(* IEC 61131-3 sources: s7-to-codesys/tests/POUs/Scenarios/FB_PumpAlternation_ScenarioTest, 7 files *)

(* ---- FB_PumpAlternation_ScenarioTest.decl.st ---- *)
// AUTO-GENERATED — не редактировать: s7conv gen-tests, сценарии scenarios/FB_PumpAlternation.csv
// Правка — в CSV (scenarios/README.md), затем python -m s7conv build-corpus.
// Назначение: тесты поведения сконвертированного FB_PumpAlternation по сценариям CSV (сценариев: 6, строк: 31):
//             один метод-тест на сценарий, строки — по порядку с моделируемым временем GVL_S7Clock.
//             Ожидаемые значения — из CSV (эталонные модели по описанию логики блока), не из
//             результата конвертации.
// Автор:      s7conv 0.1.0 (сгенерировано)
// Версия:     не указана
// Документ:   scenarios/README.md, docs/methodology.md, раздел «Проверка поведения»
FUNCTION_BLOCK FB_PumpAlternation_ScenarioTest EXTENDS coUnit.FB_TestSuite
VAR
    fbRotateOnStop : FB_PumpAlternation;  // свой экземпляр на сценарий
    xRotateOnStopDone : BOOL;  // сценарий выполнен (выполняется один раз)
    fbStandbyTakesOver : FB_PumpAlternation;  // свой экземпляр на сценарий
    xStandbyTakesOverDone : BOOL;  // сценарий выполнен (выполняется один раз)
    fbForcedAlternate : FB_PumpAlternation;  // свой экземпляр на сценарий
    xForcedAlternateDone : BOOL;  // сценарий выполнен (выполняется один раз)
    fbRotateOnStopDisabled : FB_PumpAlternation;  // свой экземпляр на сценарий
    xRotateOnStopDisabledDone : BOOL;  // сценарий выполнен (выполняется один раз)
    fbNoPumpsAvailable : FB_PumpAlternation;  // свой экземпляр на сценарий
    xNoPumpsAvailableDone : BOOL;  // сценарий выполнен (выполняется один раз)
    fbDemandClamped : FB_PumpAlternation;  // свой экземпляр на сценарий
    xDemandClampedDone : BOOL;  // сценарий выполнен (выполняется один раз)
END_VAR

(* ---- DemandClamped.method.impl.st ---- *)
// AUTO-GENERATED — не редактировать: scenarios/FB_PumpAlternation.csv, сценарий DemandClamped
coUnit.TEST('DemandClamped');
IF NOT xDemandClampedDone THEN
    xDemandClampedDone := TRUE;
    GVL_S7Clock.xSimulation := TRUE;

    // #1, t = 0 мс — demand 5 -> 3: все три
    GVL_S7Clock.tSimNow := T#0MS;
    fbDemandClamped.demand := 5;
    fbDemandClamped.available1 := TRUE;
    fbDemandClamped.available2 := TRUE;
    fbDemandClamped.available3 := TRUE;
    fbDemandClamped.alternate := FALSE;
    fbDemandClamped.rotateOnStop := TRUE;
    fbDemandClamped();
    AssertEquals_BOOL(Expected := TRUE, Actual := fbDemandClamped.run1, Message := 'DemandClamped#1 run1');
    AssertEquals_BOOL(Expected := TRUE, Actual := fbDemandClamped.run2, Message := 'DemandClamped#1 run2');
    AssertEquals_BOOL(Expected := TRUE, Actual := fbDemandClamped.run3, Message := 'DemandClamped#1 run3');
    AssertEquals_INT(Expected := 1, Actual := fbDemandClamped.leadPump, Message := 'DemandClamped#1 leadPump');
    AssertEquals_INT(Expected := 3, Actual := fbDemandClamped.runningCount, Message := 'DemandClamped#1 runningCount');
    AssertEquals_BOOL(Expected := FALSE, Actual := fbDemandClamped.shortage, Message := 'DemandClamped#1 shortage');

    // #2, t = 100 мс — demand -1 -> 0: останов, ведущий -> 2
    GVL_S7Clock.tSimNow := T#100MS;
    fbDemandClamped.demand := -1;
    fbDemandClamped();
    AssertEquals_BOOL(Expected := FALSE, Actual := fbDemandClamped.run1, Message := 'DemandClamped#2 run1');
    AssertEquals_BOOL(Expected := FALSE, Actual := fbDemandClamped.run2, Message := 'DemandClamped#2 run2');
    AssertEquals_BOOL(Expected := FALSE, Actual := fbDemandClamped.run3, Message := 'DemandClamped#2 run3');
    AssertEquals_INT(Expected := 2, Actual := fbDemandClamped.leadPump, Message := 'DemandClamped#2 leadPump');
    AssertEquals_INT(Expected := 0, Actual := fbDemandClamped.runningCount, Message := 'DemandClamped#2 runningCount');
    AssertEquals_BOOL(Expected := FALSE, Actual := fbDemandClamped.shortage, Message := 'DemandClamped#2 shortage');

    // #3, t = 200 мс — demand 4 -> 3: 2, 3, 1
    GVL_S7Clock.tSimNow := T#200MS;
    fbDemandClamped.demand := 4;
    fbDemandClamped();
    AssertEquals_BOOL(Expected := TRUE, Actual := fbDemandClamped.run1, Message := 'DemandClamped#3 run1');
    AssertEquals_BOOL(Expected := TRUE, Actual := fbDemandClamped.run2, Message := 'DemandClamped#3 run2');
    AssertEquals_BOOL(Expected := TRUE, Actual := fbDemandClamped.run3, Message := 'DemandClamped#3 run3');
    AssertEquals_INT(Expected := 2, Actual := fbDemandClamped.leadPump, Message := 'DemandClamped#3 leadPump');
    AssertEquals_INT(Expected := 3, Actual := fbDemandClamped.runningCount, Message := 'DemandClamped#3 runningCount');
    AssertEquals_BOOL(Expected := FALSE, Actual := fbDemandClamped.shortage, Message := 'DemandClamped#3 shortage');

    GVL_S7Clock.xSimulation := FALSE;
END_IF
coUnit.TEST_FINISHED();

(* ---- ForcedAlternate.method.impl.st ---- *)
// AUTO-GENERATED — не редактировать: scenarios/FB_PumpAlternation.csv, сценарий ForcedAlternate
coUnit.TEST('ForcedAlternate');
IF NOT xForcedAlternateDone THEN
    xForcedAlternateDone := TRUE;
    GVL_S7Clock.xSimulation := TRUE;

    // #1, t = 0 мс — один насос: 1
    GVL_S7Clock.tSimNow := T#0MS;
    fbForcedAlternate.demand := 1;
    fbForcedAlternate.available1 := TRUE;
    fbForcedAlternate.available2 := TRUE;
    fbForcedAlternate.available3 := TRUE;
    fbForcedAlternate.alternate := FALSE;
    fbForcedAlternate.rotateOnStop := TRUE;
    fbForcedAlternate();
    AssertEquals_BOOL(Expected := TRUE, Actual := fbForcedAlternate.run1, Message := 'ForcedAlternate#1 run1');
    AssertEquals_BOOL(Expected := FALSE, Actual := fbForcedAlternate.run2, Message := 'ForcedAlternate#1 run2');
    AssertEquals_BOOL(Expected := FALSE, Actual := fbForcedAlternate.run3, Message := 'ForcedAlternate#1 run3');
    AssertEquals_INT(Expected := 1, Actual := fbForcedAlternate.leadPump, Message := 'ForcedAlternate#1 leadPump');
    AssertEquals_INT(Expected := 1,
                     Actual := fbForcedAlternate.runningCount,
                     Message := 'ForcedAlternate#1 runningCount');
    AssertEquals_BOOL(Expected := FALSE, Actual := fbForcedAlternate.shortage, Message := 'ForcedAlternate#1 shortage');

    // #2, t = 100 мс — фронт alternate: ведущий 2, переключение в работе
    GVL_S7Clock.tSimNow := T#100MS;
    fbForcedAlternate.alternate := TRUE;
    fbForcedAlternate();
    AssertEquals_BOOL(Expected := FALSE, Actual := fbForcedAlternate.run1, Message := 'ForcedAlternate#2 run1');
    AssertEquals_BOOL(Expected := TRUE, Actual := fbForcedAlternate.run2, Message := 'ForcedAlternate#2 run2');
    AssertEquals_BOOL(Expected := FALSE, Actual := fbForcedAlternate.run3, Message := 'ForcedAlternate#2 run3');
    AssertEquals_INT(Expected := 2, Actual := fbForcedAlternate.leadPump, Message := 'ForcedAlternate#2 leadPump');
    AssertEquals_INT(Expected := 1,
                     Actual := fbForcedAlternate.runningCount,
                     Message := 'ForcedAlternate#2 runningCount');
    AssertEquals_BOOL(Expected := FALSE, Actual := fbForcedAlternate.shortage, Message := 'ForcedAlternate#2 shortage');

    // #3, t = 200 мс — alternate держится: фронта нет
    GVL_S7Clock.tSimNow := T#200MS;
    fbForcedAlternate();
    AssertEquals_BOOL(Expected := FALSE, Actual := fbForcedAlternate.run1, Message := 'ForcedAlternate#3 run1');
    AssertEquals_BOOL(Expected := TRUE, Actual := fbForcedAlternate.run2, Message := 'ForcedAlternate#3 run2');
    AssertEquals_BOOL(Expected := FALSE, Actual := fbForcedAlternate.run3, Message := 'ForcedAlternate#3 run3');
    AssertEquals_INT(Expected := 2, Actual := fbForcedAlternate.leadPump, Message := 'ForcedAlternate#3 leadPump');
    AssertEquals_INT(Expected := 1,
                     Actual := fbForcedAlternate.runningCount,
                     Message := 'ForcedAlternate#3 runningCount');
    AssertEquals_BOOL(Expected := FALSE, Actual := fbForcedAlternate.shortage, Message := 'ForcedAlternate#3 shortage');

    // #4, t = 300 мс — отпущен
    GVL_S7Clock.tSimNow := T#300MS;
    fbForcedAlternate.alternate := FALSE;
    fbForcedAlternate();
    AssertEquals_BOOL(Expected := FALSE, Actual := fbForcedAlternate.run1, Message := 'ForcedAlternate#4 run1');
    AssertEquals_BOOL(Expected := TRUE, Actual := fbForcedAlternate.run2, Message := 'ForcedAlternate#4 run2');
    AssertEquals_BOOL(Expected := FALSE, Actual := fbForcedAlternate.run3, Message := 'ForcedAlternate#4 run3');
    AssertEquals_INT(Expected := 2, Actual := fbForcedAlternate.leadPump, Message := 'ForcedAlternate#4 leadPump');
    AssertEquals_INT(Expected := 1,
                     Actual := fbForcedAlternate.runningCount,
                     Message := 'ForcedAlternate#4 runningCount');
    AssertEquals_BOOL(Expected := FALSE, Actual := fbForcedAlternate.shortage, Message := 'ForcedAlternate#4 shortage');

    // #5, t = 400 мс — фронт: ведущий 3
    GVL_S7Clock.tSimNow := T#400MS;
    fbForcedAlternate.alternate := TRUE;
    fbForcedAlternate();
    AssertEquals_BOOL(Expected := FALSE, Actual := fbForcedAlternate.run1, Message := 'ForcedAlternate#5 run1');
    AssertEquals_BOOL(Expected := FALSE, Actual := fbForcedAlternate.run2, Message := 'ForcedAlternate#5 run2');
    AssertEquals_BOOL(Expected := TRUE, Actual := fbForcedAlternate.run3, Message := 'ForcedAlternate#5 run3');
    AssertEquals_INT(Expected := 3, Actual := fbForcedAlternate.leadPump, Message := 'ForcedAlternate#5 leadPump');
    AssertEquals_INT(Expected := 1,
                     Actual := fbForcedAlternate.runningCount,
                     Message := 'ForcedAlternate#5 runningCount');
    AssertEquals_BOOL(Expected := FALSE, Actual := fbForcedAlternate.shortage, Message := 'ForcedAlternate#5 shortage');

    GVL_S7Clock.xSimulation := FALSE;
END_IF
coUnit.TEST_FINISHED();

(* ---- NoPumpsAvailable.method.impl.st ---- *)
// AUTO-GENERATED — не редактировать: scenarios/FB_PumpAlternation.csv, сценарий NoPumpsAvailable
coUnit.TEST('NoPumpsAvailable');
IF NOT xNoPumpsAvailableDone THEN
    xNoPumpsAvailableDone := TRUE;
    GVL_S7Clock.xSimulation := TRUE;

    // #1, t = 0 мс — нужно 2, доступных нет: нехватка
    GVL_S7Clock.tSimNow := T#0MS;
    fbNoPumpsAvailable.demand := 2;
    fbNoPumpsAvailable.available1 := FALSE;
    fbNoPumpsAvailable.available2 := FALSE;
    fbNoPumpsAvailable.available3 := FALSE;
    fbNoPumpsAvailable.alternate := FALSE;
    fbNoPumpsAvailable.rotateOnStop := TRUE;
    fbNoPumpsAvailable();
    AssertEquals_BOOL(Expected := FALSE, Actual := fbNoPumpsAvailable.run1, Message := 'NoPumpsAvailable#1 run1');
    AssertEquals_BOOL(Expected := FALSE, Actual := fbNoPumpsAvailable.run2, Message := 'NoPumpsAvailable#1 run2');
    AssertEquals_BOOL(Expected := FALSE, Actual := fbNoPumpsAvailable.run3, Message := 'NoPumpsAvailable#1 run3');
    AssertEquals_INT(Expected := 1, Actual := fbNoPumpsAvailable.leadPump, Message := 'NoPumpsAvailable#1 leadPump');
    AssertEquals_INT(Expected := 0,
                     Actual := fbNoPumpsAvailable.runningCount,
                     Message := 'NoPumpsAvailable#1 runningCount');
    AssertEquals_BOOL(Expected := TRUE,
                      Actual := fbNoPumpsAvailable.shortage,
                      Message := 'NoPumpsAvailable#1 shortage');

    // #2, t = 100 мс — останов: искать некого, ведущий 1
    GVL_S7Clock.tSimNow := T#100MS;
    fbNoPumpsAvailable.demand := 0;
    fbNoPumpsAvailable();
    AssertEquals_BOOL(Expected := FALSE, Actual := fbNoPumpsAvailable.run1, Message := 'NoPumpsAvailable#2 run1');
    AssertEquals_BOOL(Expected := FALSE, Actual := fbNoPumpsAvailable.run2, Message := 'NoPumpsAvailable#2 run2');
    AssertEquals_BOOL(Expected := FALSE, Actual := fbNoPumpsAvailable.run3, Message := 'NoPumpsAvailable#2 run3');
    AssertEquals_INT(Expected := 1, Actual := fbNoPumpsAvailable.leadPump, Message := 'NoPumpsAvailable#2 leadPump');
    AssertEquals_INT(Expected := 0,
                     Actual := fbNoPumpsAvailable.runningCount,
                     Message := 'NoPumpsAvailable#2 runningCount');
    AssertEquals_BOOL(Expected := FALSE,
                      Actual := fbNoPumpsAvailable.shortage,
                      Message := 'NoPumpsAvailable#2 shortage');

    // #3, t = 200 мс — фронт alternate: искать некого, ведущий 1
    GVL_S7Clock.tSimNow := T#200MS;
    fbNoPumpsAvailable.alternate := TRUE;
    fbNoPumpsAvailable();
    AssertEquals_BOOL(Expected := FALSE, Actual := fbNoPumpsAvailable.run1, Message := 'NoPumpsAvailable#3 run1');
    AssertEquals_BOOL(Expected := FALSE, Actual := fbNoPumpsAvailable.run2, Message := 'NoPumpsAvailable#3 run2');
    AssertEquals_BOOL(Expected := FALSE, Actual := fbNoPumpsAvailable.run3, Message := 'NoPumpsAvailable#3 run3');
    AssertEquals_INT(Expected := 1, Actual := fbNoPumpsAvailable.leadPump, Message := 'NoPumpsAvailable#3 leadPump');
    AssertEquals_INT(Expected := 0,
                     Actual := fbNoPumpsAvailable.runningCount,
                     Message := 'NoPumpsAvailable#3 runningCount');
    AssertEquals_BOOL(Expected := FALSE,
                      Actual := fbNoPumpsAvailable.shortage,
                      Message := 'NoPumpsAvailable#3 shortage');

    // #4, t = 300 мс — доступен только 3: работает 3, ведущий 1
    GVL_S7Clock.tSimNow := T#300MS;
    fbNoPumpsAvailable.demand := 1;
    fbNoPumpsAvailable.available3 := TRUE;
    fbNoPumpsAvailable.alternate := FALSE;
    fbNoPumpsAvailable();
    AssertEquals_BOOL(Expected := FALSE, Actual := fbNoPumpsAvailable.run1, Message := 'NoPumpsAvailable#4 run1');
    AssertEquals_BOOL(Expected := FALSE, Actual := fbNoPumpsAvailable.run2, Message := 'NoPumpsAvailable#4 run2');
    AssertEquals_BOOL(Expected := TRUE, Actual := fbNoPumpsAvailable.run3, Message := 'NoPumpsAvailable#4 run3');
    AssertEquals_INT(Expected := 1, Actual := fbNoPumpsAvailable.leadPump, Message := 'NoPumpsAvailable#4 leadPump');
    AssertEquals_INT(Expected := 1,
                     Actual := fbNoPumpsAvailable.runningCount,
                     Message := 'NoPumpsAvailable#4 runningCount');
    AssertEquals_BOOL(Expected := FALSE,
                      Actual := fbNoPumpsAvailable.shortage,
                      Message := 'NoPumpsAvailable#4 shortage');

    GVL_S7Clock.xSimulation := FALSE;
END_IF
coUnit.TEST_FINISHED();

(* ---- RotateOnStop.method.impl.st ---- *)
// AUTO-GENERATED — не редактировать: scenarios/FB_PumpAlternation.csv, сценарий RotateOnStop
coUnit.TEST('RotateOnStop');
IF NOT xRotateOnStopDone THEN
    xRotateOnStopDone := TRUE;
    GVL_S7Clock.xSimulation := TRUE;

    // #1, t = 0 мс — первый вызов при demand = 0: спада нет, ведущий 1
    GVL_S7Clock.tSimNow := T#0MS;
    fbRotateOnStop.demand := 0;
    fbRotateOnStop.available1 := TRUE;
    fbRotateOnStop.available2 := TRUE;
    fbRotateOnStop.available3 := TRUE;
    fbRotateOnStop.alternate := FALSE;
    fbRotateOnStop.rotateOnStop := TRUE;
    fbRotateOnStop();
    AssertEquals_BOOL(Expected := FALSE, Actual := fbRotateOnStop.run1, Message := 'RotateOnStop#1 run1');
    AssertEquals_BOOL(Expected := FALSE, Actual := fbRotateOnStop.run2, Message := 'RotateOnStop#1 run2');
    AssertEquals_BOOL(Expected := FALSE, Actual := fbRotateOnStop.run3, Message := 'RotateOnStop#1 run3');
    AssertEquals_INT(Expected := 1, Actual := fbRotateOnStop.leadPump, Message := 'RotateOnStop#1 leadPump');
    AssertEquals_INT(Expected := 0, Actual := fbRotateOnStop.runningCount, Message := 'RotateOnStop#1 runningCount');
    AssertEquals_BOOL(Expected := FALSE, Actual := fbRotateOnStop.shortage, Message := 'RotateOnStop#1 shortage');

    // #2, t = 100 мс — один насос: ведущий 1
    GVL_S7Clock.tSimNow := T#100MS;
    fbRotateOnStop.demand := 1;
    fbRotateOnStop();
    AssertEquals_BOOL(Expected := TRUE, Actual := fbRotateOnStop.run1, Message := 'RotateOnStop#2 run1');
    AssertEquals_BOOL(Expected := FALSE, Actual := fbRotateOnStop.run2, Message := 'RotateOnStop#2 run2');
    AssertEquals_BOOL(Expected := FALSE, Actual := fbRotateOnStop.run3, Message := 'RotateOnStop#2 run3');
    AssertEquals_INT(Expected := 1, Actual := fbRotateOnStop.leadPump, Message := 'RotateOnStop#2 leadPump');
    AssertEquals_INT(Expected := 1, Actual := fbRotateOnStop.runningCount, Message := 'RotateOnStop#2 runningCount');
    AssertEquals_BOOL(Expected := FALSE, Actual := fbRotateOnStop.shortage, Message := 'RotateOnStop#2 shortage');

    // #3, t = 200 мс — два насоса: 1 и 2
    GVL_S7Clock.tSimNow := T#200MS;
    fbRotateOnStop.demand := 2;
    fbRotateOnStop();
    AssertEquals_BOOL(Expected := TRUE, Actual := fbRotateOnStop.run1, Message := 'RotateOnStop#3 run1');
    AssertEquals_BOOL(Expected := TRUE, Actual := fbRotateOnStop.run2, Message := 'RotateOnStop#3 run2');
    AssertEquals_BOOL(Expected := FALSE, Actual := fbRotateOnStop.run3, Message := 'RotateOnStop#3 run3');
    AssertEquals_INT(Expected := 1, Actual := fbRotateOnStop.leadPump, Message := 'RotateOnStop#3 leadPump');
    AssertEquals_INT(Expected := 2, Actual := fbRotateOnStop.runningCount, Message := 'RotateOnStop#3 runningCount');
    AssertEquals_BOOL(Expected := FALSE, Actual := fbRotateOnStop.shortage, Message := 'RotateOnStop#3 shortage');

    // #4, t = 300 мс — останов группы: ведущий -> 2
    GVL_S7Clock.tSimNow := T#300MS;
    fbRotateOnStop.demand := 0;
    fbRotateOnStop();
    AssertEquals_BOOL(Expected := FALSE, Actual := fbRotateOnStop.run1, Message := 'RotateOnStop#4 run1');
    AssertEquals_BOOL(Expected := FALSE, Actual := fbRotateOnStop.run2, Message := 'RotateOnStop#4 run2');
    AssertEquals_BOOL(Expected := FALSE, Actual := fbRotateOnStop.run3, Message := 'RotateOnStop#4 run3');
    AssertEquals_INT(Expected := 2, Actual := fbRotateOnStop.leadPump, Message := 'RotateOnStop#4 leadPump');
    AssertEquals_INT(Expected := 0, Actual := fbRotateOnStop.runningCount, Message := 'RotateOnStop#4 runningCount');
    AssertEquals_BOOL(Expected := FALSE, Actual := fbRotateOnStop.shortage, Message := 'RotateOnStop#4 shortage');

    // #5, t = 400 мс — один насос: 2
    GVL_S7Clock.tSimNow := T#400MS;
    fbRotateOnStop.demand := 1;
    fbRotateOnStop();
    AssertEquals_BOOL(Expected := FALSE, Actual := fbRotateOnStop.run1, Message := 'RotateOnStop#5 run1');
    AssertEquals_BOOL(Expected := TRUE, Actual := fbRotateOnStop.run2, Message := 'RotateOnStop#5 run2');
    AssertEquals_BOOL(Expected := FALSE, Actual := fbRotateOnStop.run3, Message := 'RotateOnStop#5 run3');
    AssertEquals_INT(Expected := 2, Actual := fbRotateOnStop.leadPump, Message := 'RotateOnStop#5 leadPump');
    AssertEquals_INT(Expected := 1, Actual := fbRotateOnStop.runningCount, Message := 'RotateOnStop#5 runningCount');
    AssertEquals_BOOL(Expected := FALSE, Actual := fbRotateOnStop.shortage, Message := 'RotateOnStop#5 shortage');

    // #6, t = 500 мс — три насоса: 2, 3, 1
    GVL_S7Clock.tSimNow := T#500MS;
    fbRotateOnStop.demand := 3;
    fbRotateOnStop();
    AssertEquals_BOOL(Expected := TRUE, Actual := fbRotateOnStop.run1, Message := 'RotateOnStop#6 run1');
    AssertEquals_BOOL(Expected := TRUE, Actual := fbRotateOnStop.run2, Message := 'RotateOnStop#6 run2');
    AssertEquals_BOOL(Expected := TRUE, Actual := fbRotateOnStop.run3, Message := 'RotateOnStop#6 run3');
    AssertEquals_INT(Expected := 2, Actual := fbRotateOnStop.leadPump, Message := 'RotateOnStop#6 leadPump');
    AssertEquals_INT(Expected := 3, Actual := fbRotateOnStop.runningCount, Message := 'RotateOnStop#6 runningCount');
    AssertEquals_BOOL(Expected := FALSE, Actual := fbRotateOnStop.shortage, Message := 'RotateOnStop#6 shortage');

    // #7, t = 600 мс — останов: ведущий -> 3
    GVL_S7Clock.tSimNow := T#600MS;
    fbRotateOnStop.demand := 0;
    fbRotateOnStop();
    AssertEquals_BOOL(Expected := FALSE, Actual := fbRotateOnStop.run1, Message := 'RotateOnStop#7 run1');
    AssertEquals_BOOL(Expected := FALSE, Actual := fbRotateOnStop.run2, Message := 'RotateOnStop#7 run2');
    AssertEquals_BOOL(Expected := FALSE, Actual := fbRotateOnStop.run3, Message := 'RotateOnStop#7 run3');
    AssertEquals_INT(Expected := 3, Actual := fbRotateOnStop.leadPump, Message := 'RotateOnStop#7 leadPump');
    AssertEquals_INT(Expected := 0, Actual := fbRotateOnStop.runningCount, Message := 'RotateOnStop#7 runningCount');
    AssertEquals_BOOL(Expected := FALSE, Actual := fbRotateOnStop.shortage, Message := 'RotateOnStop#7 shortage');

    // #8, t = 700 мс — один насос: 3
    GVL_S7Clock.tSimNow := T#700MS;
    fbRotateOnStop.demand := 1;
    fbRotateOnStop();
    AssertEquals_BOOL(Expected := FALSE, Actual := fbRotateOnStop.run1, Message := 'RotateOnStop#8 run1');
    AssertEquals_BOOL(Expected := FALSE, Actual := fbRotateOnStop.run2, Message := 'RotateOnStop#8 run2');
    AssertEquals_BOOL(Expected := TRUE, Actual := fbRotateOnStop.run3, Message := 'RotateOnStop#8 run3');
    AssertEquals_INT(Expected := 3, Actual := fbRotateOnStop.leadPump, Message := 'RotateOnStop#8 leadPump');
    AssertEquals_INT(Expected := 1, Actual := fbRotateOnStop.runningCount, Message := 'RotateOnStop#8 runningCount');
    AssertEquals_BOOL(Expected := FALSE, Actual := fbRotateOnStop.shortage, Message := 'RotateOnStop#8 shortage');

    // #9, t = 800 мс — останов: ведущий -> 1 (по кругу)
    GVL_S7Clock.tSimNow := T#800MS;
    fbRotateOnStop.demand := 0;
    fbRotateOnStop();
    AssertEquals_BOOL(Expected := FALSE, Actual := fbRotateOnStop.run1, Message := 'RotateOnStop#9 run1');
    AssertEquals_BOOL(Expected := FALSE, Actual := fbRotateOnStop.run2, Message := 'RotateOnStop#9 run2');
    AssertEquals_BOOL(Expected := FALSE, Actual := fbRotateOnStop.run3, Message := 'RotateOnStop#9 run3');
    AssertEquals_INT(Expected := 1, Actual := fbRotateOnStop.leadPump, Message := 'RotateOnStop#9 leadPump');
    AssertEquals_INT(Expected := 0, Actual := fbRotateOnStop.runningCount, Message := 'RotateOnStop#9 runningCount');
    AssertEquals_BOOL(Expected := FALSE, Actual := fbRotateOnStop.shortage, Message := 'RotateOnStop#9 shortage');

    // #10, t = 900 мс — demand остаётся 0: спада нет, ведущий 1
    GVL_S7Clock.tSimNow := T#900MS;
    fbRotateOnStop();
    AssertEquals_BOOL(Expected := FALSE, Actual := fbRotateOnStop.run1, Message := 'RotateOnStop#10 run1');
    AssertEquals_BOOL(Expected := FALSE, Actual := fbRotateOnStop.run2, Message := 'RotateOnStop#10 run2');
    AssertEquals_BOOL(Expected := FALSE, Actual := fbRotateOnStop.run3, Message := 'RotateOnStop#10 run3');
    AssertEquals_INT(Expected := 1, Actual := fbRotateOnStop.leadPump, Message := 'RotateOnStop#10 leadPump');
    AssertEquals_INT(Expected := 0, Actual := fbRotateOnStop.runningCount, Message := 'RotateOnStop#10 runningCount');
    AssertEquals_BOOL(Expected := FALSE, Actual := fbRotateOnStop.shortage, Message := 'RotateOnStop#10 shortage');

    GVL_S7Clock.xSimulation := FALSE;
END_IF
coUnit.TEST_FINISHED();

(* ---- RotateOnStopDisabled.method.impl.st ---- *)
// AUTO-GENERATED — не редактировать: scenarios/FB_PumpAlternation.csv, сценарий RotateOnStopDisabled
coUnit.TEST('RotateOnStopDisabled');
IF NOT xRotateOnStopDisabledDone THEN
    xRotateOnStopDisabledDone := TRUE;
    GVL_S7Clock.xSimulation := TRUE;

    // #1, t = 0 мс — один насос: 1
    GVL_S7Clock.tSimNow := T#0MS;
    fbRotateOnStopDisabled.demand := 1;
    fbRotateOnStopDisabled.available1 := TRUE;
    fbRotateOnStopDisabled.available2 := TRUE;
    fbRotateOnStopDisabled.available3 := TRUE;
    fbRotateOnStopDisabled.alternate := FALSE;
    fbRotateOnStopDisabled.rotateOnStop := FALSE;
    fbRotateOnStopDisabled();
    AssertEquals_BOOL(Expected := TRUE,
                      Actual := fbRotateOnStopDisabled.run1,
                      Message := 'RotateOnStopDisabled#1 run1');
    AssertEquals_BOOL(Expected := FALSE,
                      Actual := fbRotateOnStopDisabled.run2,
                      Message := 'RotateOnStopDisabled#1 run2');
    AssertEquals_BOOL(Expected := FALSE,
                      Actual := fbRotateOnStopDisabled.run3,
                      Message := 'RotateOnStopDisabled#1 run3');
    AssertEquals_INT(Expected := 1,
                     Actual := fbRotateOnStopDisabled.leadPump,
                     Message := 'RotateOnStopDisabled#1 leadPump');
    AssertEquals_INT(Expected := 1,
                     Actual := fbRotateOnStopDisabled.runningCount,
                     Message := 'RotateOnStopDisabled#1 runningCount');
    AssertEquals_BOOL(Expected := FALSE,
                      Actual := fbRotateOnStopDisabled.shortage,
                      Message := 'RotateOnStopDisabled#1 shortage');

    // #2, t = 100 мс — останов: ведущий остаётся 1
    GVL_S7Clock.tSimNow := T#100MS;
    fbRotateOnStopDisabled.demand := 0;
    fbRotateOnStopDisabled();
    AssertEquals_BOOL(Expected := FALSE,
                      Actual := fbRotateOnStopDisabled.run1,
                      Message := 'RotateOnStopDisabled#2 run1');
    AssertEquals_BOOL(Expected := FALSE,
                      Actual := fbRotateOnStopDisabled.run2,
                      Message := 'RotateOnStopDisabled#2 run2');
    AssertEquals_BOOL(Expected := FALSE,
                      Actual := fbRotateOnStopDisabled.run3,
                      Message := 'RotateOnStopDisabled#2 run3');
    AssertEquals_INT(Expected := 1,
                     Actual := fbRotateOnStopDisabled.leadPump,
                     Message := 'RotateOnStopDisabled#2 leadPump');
    AssertEquals_INT(Expected := 0,
                     Actual := fbRotateOnStopDisabled.runningCount,
                     Message := 'RotateOnStopDisabled#2 runningCount');
    AssertEquals_BOOL(Expected := FALSE,
                      Actual := fbRotateOnStopDisabled.shortage,
                      Message := 'RotateOnStopDisabled#2 shortage');

    // #3, t = 200 мс — снова 1
    GVL_S7Clock.tSimNow := T#200MS;
    fbRotateOnStopDisabled.demand := 1;
    fbRotateOnStopDisabled();
    AssertEquals_BOOL(Expected := TRUE,
                      Actual := fbRotateOnStopDisabled.run1,
                      Message := 'RotateOnStopDisabled#3 run1');
    AssertEquals_BOOL(Expected := FALSE,
                      Actual := fbRotateOnStopDisabled.run2,
                      Message := 'RotateOnStopDisabled#3 run2');
    AssertEquals_BOOL(Expected := FALSE,
                      Actual := fbRotateOnStopDisabled.run3,
                      Message := 'RotateOnStopDisabled#3 run3');
    AssertEquals_INT(Expected := 1,
                     Actual := fbRotateOnStopDisabled.leadPump,
                     Message := 'RotateOnStopDisabled#3 leadPump');
    AssertEquals_INT(Expected := 1,
                     Actual := fbRotateOnStopDisabled.runningCount,
                     Message := 'RotateOnStopDisabled#3 runningCount');
    AssertEquals_BOOL(Expected := FALSE,
                      Actual := fbRotateOnStopDisabled.shortage,
                      Message := 'RotateOnStopDisabled#3 shortage');

    GVL_S7Clock.xSimulation := FALSE;
END_IF
coUnit.TEST_FINISHED();

(* ---- StandbyTakesOver.method.impl.st ---- *)
// AUTO-GENERATED — не редактировать: scenarios/FB_PumpAlternation.csv, сценарий StandbyTakesOver
coUnit.TEST('StandbyTakesOver');
IF NOT xStandbyTakesOverDone THEN
    xStandbyTakesOverDone := TRUE;
    GVL_S7Clock.xSimulation := TRUE;

    // #1, t = 0 мс — один насос: 1
    GVL_S7Clock.tSimNow := T#0MS;
    fbStandbyTakesOver.demand := 1;
    fbStandbyTakesOver.available1 := TRUE;
    fbStandbyTakesOver.available2 := TRUE;
    fbStandbyTakesOver.available3 := TRUE;
    fbStandbyTakesOver.alternate := FALSE;
    fbStandbyTakesOver.rotateOnStop := TRUE;
    fbStandbyTakesOver();
    AssertEquals_BOOL(Expected := TRUE, Actual := fbStandbyTakesOver.run1, Message := 'StandbyTakesOver#1 run1');
    AssertEquals_BOOL(Expected := FALSE, Actual := fbStandbyTakesOver.run2, Message := 'StandbyTakesOver#1 run2');
    AssertEquals_BOOL(Expected := FALSE, Actual := fbStandbyTakesOver.run3, Message := 'StandbyTakesOver#1 run3');
    AssertEquals_INT(Expected := 1, Actual := fbStandbyTakesOver.leadPump, Message := 'StandbyTakesOver#1 leadPump');
    AssertEquals_INT(Expected := 1,
                     Actual := fbStandbyTakesOver.runningCount,
                     Message := 'StandbyTakesOver#1 runningCount');
    AssertEquals_BOOL(Expected := FALSE,
                      Actual := fbStandbyTakesOver.shortage,
                      Message := 'StandbyTakesOver#1 shortage');

    // #2, t = 100 мс — насос 1 недоступен: работает 2, ведущий остаётся 1
    GVL_S7Clock.tSimNow := T#100MS;
    fbStandbyTakesOver.available1 := FALSE;
    fbStandbyTakesOver();
    AssertEquals_BOOL(Expected := FALSE, Actual := fbStandbyTakesOver.run1, Message := 'StandbyTakesOver#2 run1');
    AssertEquals_BOOL(Expected := TRUE, Actual := fbStandbyTakesOver.run2, Message := 'StandbyTakesOver#2 run2');
    AssertEquals_BOOL(Expected := FALSE, Actual := fbStandbyTakesOver.run3, Message := 'StandbyTakesOver#2 run3');
    AssertEquals_INT(Expected := 1, Actual := fbStandbyTakesOver.leadPump, Message := 'StandbyTakesOver#2 leadPump');
    AssertEquals_INT(Expected := 1,
                     Actual := fbStandbyTakesOver.runningCount,
                     Message := 'StandbyTakesOver#2 runningCount');
    AssertEquals_BOOL(Expected := FALSE,
                      Actual := fbStandbyTakesOver.shortage,
                      Message := 'StandbyTakesOver#2 shortage');

    // #3, t = 200 мс — насос 1 вернулся: снова 1
    GVL_S7Clock.tSimNow := T#200MS;
    fbStandbyTakesOver.available1 := TRUE;
    fbStandbyTakesOver();
    AssertEquals_BOOL(Expected := TRUE, Actual := fbStandbyTakesOver.run1, Message := 'StandbyTakesOver#3 run1');
    AssertEquals_BOOL(Expected := FALSE, Actual := fbStandbyTakesOver.run2, Message := 'StandbyTakesOver#3 run2');
    AssertEquals_BOOL(Expected := FALSE, Actual := fbStandbyTakesOver.run3, Message := 'StandbyTakesOver#3 run3');
    AssertEquals_INT(Expected := 1, Actual := fbStandbyTakesOver.leadPump, Message := 'StandbyTakesOver#3 leadPump');
    AssertEquals_INT(Expected := 1,
                     Actual := fbStandbyTakesOver.runningCount,
                     Message := 'StandbyTakesOver#3 runningCount');
    AssertEquals_BOOL(Expected := FALSE,
                      Actual := fbStandbyTakesOver.shortage,
                      Message := 'StandbyTakesOver#3 shortage');

    // #4, t = 300 мс — нужно 3, доступно 2: 1 и 3, нехватка
    GVL_S7Clock.tSimNow := T#300MS;
    fbStandbyTakesOver.demand := 3;
    fbStandbyTakesOver.available2 := FALSE;
    fbStandbyTakesOver();
    AssertEquals_BOOL(Expected := TRUE, Actual := fbStandbyTakesOver.run1, Message := 'StandbyTakesOver#4 run1');
    AssertEquals_BOOL(Expected := FALSE, Actual := fbStandbyTakesOver.run2, Message := 'StandbyTakesOver#4 run2');
    AssertEquals_BOOL(Expected := TRUE, Actual := fbStandbyTakesOver.run3, Message := 'StandbyTakesOver#4 run3');
    AssertEquals_INT(Expected := 1, Actual := fbStandbyTakesOver.leadPump, Message := 'StandbyTakesOver#4 leadPump');
    AssertEquals_INT(Expected := 2,
                     Actual := fbStandbyTakesOver.runningCount,
                     Message := 'StandbyTakesOver#4 runningCount');
    AssertEquals_BOOL(Expected := TRUE,
                      Actual := fbStandbyTakesOver.shortage,
                      Message := 'StandbyTakesOver#4 shortage');

    // #5, t = 400 мс — останов: после 1 недоступен 2 — ведущий 3
    GVL_S7Clock.tSimNow := T#400MS;
    fbStandbyTakesOver.demand := 0;
    fbStandbyTakesOver();
    AssertEquals_BOOL(Expected := FALSE, Actual := fbStandbyTakesOver.run1, Message := 'StandbyTakesOver#5 run1');
    AssertEquals_BOOL(Expected := FALSE, Actual := fbStandbyTakesOver.run2, Message := 'StandbyTakesOver#5 run2');
    AssertEquals_BOOL(Expected := FALSE, Actual := fbStandbyTakesOver.run3, Message := 'StandbyTakesOver#5 run3');
    AssertEquals_INT(Expected := 3, Actual := fbStandbyTakesOver.leadPump, Message := 'StandbyTakesOver#5 leadPump');
    AssertEquals_INT(Expected := 0,
                     Actual := fbStandbyTakesOver.runningCount,
                     Message := 'StandbyTakesOver#5 runningCount');
    AssertEquals_BOOL(Expected := FALSE,
                      Actual := fbStandbyTakesOver.shortage,
                      Message := 'StandbyTakesOver#5 shortage');

    // #6, t = 500 мс — один насос: 3
    GVL_S7Clock.tSimNow := T#500MS;
    fbStandbyTakesOver.demand := 1;
    fbStandbyTakesOver();
    AssertEquals_BOOL(Expected := FALSE, Actual := fbStandbyTakesOver.run1, Message := 'StandbyTakesOver#6 run1');
    AssertEquals_BOOL(Expected := FALSE, Actual := fbStandbyTakesOver.run2, Message := 'StandbyTakesOver#6 run2');
    AssertEquals_BOOL(Expected := TRUE, Actual := fbStandbyTakesOver.run3, Message := 'StandbyTakesOver#6 run3');
    AssertEquals_INT(Expected := 3, Actual := fbStandbyTakesOver.leadPump, Message := 'StandbyTakesOver#6 leadPump');
    AssertEquals_INT(Expected := 1,
                     Actual := fbStandbyTakesOver.runningCount,
                     Message := 'StandbyTakesOver#6 runningCount');
    AssertEquals_BOOL(Expected := FALSE,
                      Actual := fbStandbyTakesOver.shortage,
                      Message := 'StandbyTakesOver#6 shortage');

    GVL_S7Clock.xSimulation := FALSE;
END_IF
coUnit.TEST_FINISHED();
